{attribute 'qualified_only'}
{attribute 'strict'}
{attribute 'to_string'}
TYPE E_ModeZone :
(
	eNone := 0,
	eMain,
	
	eCIP,
	eTank1,(*Tank*)
	eTank2,(*Tank*)
	eTank3,(*Tank*)
	eTank4,(*Tank*)
	
	eProduction_Marinade,(*Line*)
	eProduction_Color,(*Line*)
	
	eTriBlender_Marinade,(*Line*)
	eTriBlender_Color,(*Line*)
	eWater,(*Line*)
	eHotWater,(*Line*)
	eLast
);
END_TYPE

(* stored: Version 1.1.0.1, ProductVersion 3.1.4024.13
   DUT E_ModeZone: Id {efef26dd-c16b-43e4-b551-d6791a077621} *)
